Fanuc KAREL source: ka00056.KL

-- PROVISIONAL review KL for V770-1; original PC SHA256 dbb2149f5ad215961a863b865db83f70ed8a74a8a1e5e3772f16c1aca833eb0d
-- Incomplete behavior may be omitted. Consult companion uncertainty JSON. Do not deploy.
PROGRAM KA00056
%NOLOCKGROUP
-- UNRESOLVED_DECL SRC type=000101
-- UNRESOLVED_DECL DST type=000199
BEGIN
  -- UNRESOLVED_PC offsets 5-25; opcodes 49,7E,4A
  -- UNRESOLVED_PC offsets 30-34; opcodes 7F
END KA00056
